Fanuc KAREL source: KA00222.KL

PROGRAM KA00222
%NOLOCKGROUP
VAR
  SRC: ARRAY[4] OF JOINTPOS
  DST: ARRAY[4] OF SHORT
BEGIN
  DST = SRC
END KA00222
